Fanuc KAREL source: KC00003.KL

PROGRAM KC00003
%NOLOCKGROUP
%ENVIRONMENT PC
VAR
  I: INTEGER
  J: INTEGER
  K: INTEGER
  R: REAL
  B: BOOLEAN
  S: STRING[80]
  T: STRING[80]
  P: PATH
  Q: PATH
  AI: ARRAY[8] OF INTEGER
  AB: ARRAY[244] OF BYTE
BEGIN
  ADD_REALPC(AB,I,R,K)
END KC00003
